(* IEC 61131-3 sources: rusty/tests/lit/multi/destructors/src, 4 files *)

(* ---- main.st ---- *)
FUNCTION main: DINT
    printf('main done$N');
END_FUNCTION

(* ---- first.st ---- *)
FUNCTION_BLOCK First
    METHOD FB_INIT
        printf('init first$N');
    END_METHOD

    METHOD FB_EXIT
        printf('exit first$N');
    END_METHOD
END_FUNCTION_BLOCK

VAR_GLOBAL
    first: First;
END_VAR

(* ---- second.st ---- *)
FUNCTION_BLOCK Second
    METHOD FB_INIT
        printf('init second$N');
    END_METHOD

    METHOD FB_EXIT
        printf('exit second$N');
    END_METHOD
END_FUNCTION_BLOCK

VAR_GLOBAL
    second: Second;
END_VAR

(* ---- third.st ---- *)
PROGRAM third
    METHOD FB_INIT
        printf('init third$N');
    END_METHOD

    METHOD FB_EXIT
        printf('exit third$N');
    END_METHOD
END_PROGRAM
